Fanuc KAREL source: KD00030.KL

PROGRAM KD00030
%NOLOCKGROUP
VAR
  I: INTEGER
  J: INTEGER
  B: BOOLEAN
  R: REAL
  S: STRING[80]
BEGIN
  CONDITION[1]:
  WHEN ABORT DO
    I = 1
  ENDCONDITION
END KD00030
